// TIA Portal V18 export
TYPE "Comm"
   STRUCT
      Connection_ID : Word;
      R_ID : CONN_R_ID;
      REQ : Bool;
      Len : Word;
      Result : Struct
         DONE : Bool;
         ERROR : Bool;
         STATUS : Word;
      END_STRUCT;
      Diagnostic : Struct
         countDone : Int;
         countError : Int;
         memStatus : Word;
      END_STRUCT;
   END_STRUCT;
END_TYPE
